// TIA Portal project "CraneSim" (V18)

(* hardware
DEVICE "S7-1500/ET200MP station_1"  S7-1500 station
   slot 0: "Rail_0"  Rack  6ES7 590-1***0-0AA0
   slot 1: "PLC_1"  CPU 1511-1 PN  6ES7 511-1AK02-0AB0  V2.9
      slot 3: "CPU display_1"  6ES7591-1AA00-0AA0
      slot 32768: "PROFINET interface_1"  X1
         slot 32769: "Port_1"  X1 P1
         slot 32770: "Port_2"  X1 P2
      slot 34817: "Virtual CP interface port_1"  Virtual CP interface port  Virtual CP interface port
*)

// ===== PLC "PLC_1"  CPU 1511-1 PN =====

VAR_GLOBAL   // PLC tag table "Default tag table"
   "Clock_Byte" AT %MB0 : Byte;
   "Clock_10Hz" AT %M0.0 : Bool;
   "Clock_5Hz" AT %M0.1 : Bool;
   "Clock_2.5Hz" AT %M0.2 : Bool;
   "Clock_2Hz" AT %M0.3 : Bool;
   "Clock_1.25Hz" AT %M0.4 : Bool;
   "Clock_1Hz" AT %M0.5 : Bool;
   "Clock_0.625Hz" AT %M0.6 : Bool;
   "Clock_0.5Hz" AT %M0.7 : Bool;
END_VAR

TYPE "typeTask"
   STRUCT
      station : Int;
      dwell_s : Int;
      crane : String[4];
      tank_name : String[10];
      prev : Int;
      next : Int;
      status : Int;
   END_STRUCT;
END_TYPE

DATA_BLOCK "Line4Data"   // DB2
{ S7_Optimized_Access := 'TRUE' }
VERSION : 0.1
   VAR
      task_count : Int;
      tasks : Array[1..20] of "typeTask";
      cmd_send : Bool;
      sts_busy : Bool;
      sts_done : Bool;
      sts_step : Int;
      sts_state : Int;
      ls_at : Array[0..9] of Bool;
      ls_dip : Bool;
      ls_up : Bool;
      btn_start : Bool;
      mv_fwd : Bool;
      mv_rev : Bool;
      mv_up : Bool;
      mv_down : Bool;
   END_VAR
BEGIN
END_DATA_BLOCK

DATA_BLOCK "CraneSequencer_DB"   // DB3
{ S7_Optimized_Access := 'TRUE' }
VERSION : 0.1
// stored: InstanceOfName CraneSequencer
"CraneSequencer"
BEGIN
END_DATA_BLOCK

FUNCTION_BLOCK "CraneSequencer"   // FB1, SCL
{ S7_Optimized_Access := 'TRUE' }
VERSION : 0.1
   VAR
      state : Int;
      idx : Int;
      count : Int;
      cur : Int;
      prevSend : Bool;
      tHold : TON_TIME;
      tDwell : TON_TIME;
   END_VAR
   VAR_TEMP
      target : Int;
      arrived : Bool;
   END_VAR
BEGIN
   // CraneSequencer — runs the Line4Data.tasks[] batch through the crane sequence.
   // Call every scan from OB1. Shared data lives in global DB "Line4Data".
   // Stations: 0=Parking 1=Loading 2..N=tanks.

   "Line4Data".sts_state := #state;

   CASE #state OF
       0:
           "Line4Data".mv_fwd := FALSE;
           "Line4Data".mv_rev := FALSE;
           "Line4Data".mv_up := FALSE;
           "Line4Data".mv_down := FALSE;
           "Line4Data".sts_busy := FALSE;
           "Line4Data".sts_step := 0;
           IF "Line4Data".cmd_send AND NOT #prevSend AND "Line4Data".task_count > 0 THEN
               #count := "Line4Data".task_count;
               #idx := 1;
               "Line4Data".sts_done := FALSE;
               "Line4Data".sts_busy := TRUE;
               #state := 10;
           END_IF;

       10:
           "Line4Data".sts_busy := TRUE;
           #target := 1;
           #arrived := "TravelTo"(target := #target, cur := #cur, atTarget := "Line4Data".ls_at[#target], fwd => "Line4Data".mv_fwd, rev => "Line4Data".mv_rev);
           IF #arrived THEN
               #cur := #target;
               "Line4Data".mv_fwd := FALSE;
               "Line4Data".mv_rev := FALSE;
               #state := 20;
           END_IF;

       20:
           "Line4Data".mv_up := FALSE;
           "Line4Data".mv_down := TRUE;
           IF "Line4Data".ls_dip THEN
               "Line4Data".mv_down := FALSE;
               #state := 30;
           END_IF;

       30:
           #tHold(IN := "Line4Data".btn_start,
                  PT := T#3S);
           IF #tHold.Q THEN
               #state := 40;
           END_IF;

       40:
           "Line4Data".mv_down := FALSE;
           "Line4Data".mv_up := TRUE;
           IF "Line4Data".ls_up THEN
               "Line4Data".mv_up := FALSE;
               #state := 50;
           END_IF;

       50:
           "Line4Data".sts_step := #idx;
           "Line4Data".tasks[#idx].status := 1;
           #target := "Line4Data".tasks[#idx].station;
           #arrived := "TravelTo"(target := #target, cur := #cur, atTarget := "Line4Data".ls_at[#target], fwd => "Line4Data".mv_fwd, rev => "Line4Data".mv_rev);
           IF #arrived THEN
               #cur := #target;
               "Line4Data".mv_fwd := FALSE;
               "Line4Data".mv_rev := FALSE;
               #state := 60;
           END_IF;

       60:
           "Line4Data".mv_up := FALSE;
           "Line4Data".mv_down := TRUE;
           IF "Line4Data".ls_dip THEN
               "Line4Data".mv_down := FALSE;
               #state := 70;
           END_IF;

       70:
           #tDwell(IN := TRUE,
                   PT := DINT_TO_TIME(INT_TO_DINT("Line4Data".tasks[#idx].dwell_s) * 1000));
           IF #tDwell.Q THEN
               #tDwell(IN := FALSE,
                       PT := T#0S);
               #state := 80;
           END_IF;

       80:
           "Line4Data".mv_down := FALSE;
           "Line4Data".mv_up := TRUE;
           IF "Line4Data".ls_up THEN
               "Line4Data".mv_up := FALSE;
               "Line4Data".tasks[#idx].status := 2;
               IF #idx < #count THEN
                   #idx := #idx + 1;
                   #state := 50;
               ELSE
                   #state := 85;
               END_IF;
           END_IF;

       85:
           #target := 0;
           #arrived := "TravelTo"(target := #target, cur := #cur, atTarget := "Line4Data".ls_at[#target], fwd => "Line4Data".mv_fwd, rev => "Line4Data".mv_rev);
           IF #arrived THEN
               #cur := #target;
               "Line4Data".mv_fwd := FALSE;
               "Line4Data".mv_rev := FALSE;
               #state := 90;
           END_IF;

       90:
           "Line4Data".sts_busy := FALSE;
           "Line4Data".sts_done := TRUE;
           IF NOT "Line4Data".cmd_send THEN
               "Line4Data".sts_done := FALSE;
               "Line4Data".sts_step := 0;
               #state := 0;
           END_IF;
   END_CASE;

   #prevSend := "Line4Data".cmd_send;
END_FUNCTION_BLOCK

FUNCTION "TravelTo" : Bool   // FC2, SCL
{ S7_Optimized_Access := 'TRUE' }
VERSION : 0.1
   VAR_INPUT
      target : Int;
      cur : Int;
      atTarget : Bool;
   END_VAR
   VAR_OUTPUT
      fwd : Bool;
      rev : Bool;
   END_VAR
BEGIN
   // TravelTo — pick the travel direction toward a target station.
   // Returns TRUE when the target limit switch is already made (arrived → stop).
   #fwd := FALSE;
   #rev := FALSE;

   IF #atTarget THEN
       ;                       // arrived: leave both motors off
   ELSIF #target > #cur THEN
       #fwd := TRUE;           // higher station number → travel forward
   ELSE
       #rev := TRUE;           // lower station number → travel reverse
   END_IF;

   #TravelTo := #atTarget;
END_FUNCTION

ORGANIZATION_BLOCK "Main"   // OB1, LAD, ProgramCycle
TITLE = "Main Program Sweep (Cycle)"
{ S7_Optimized_Access := 'TRUE' }
VERSION : 0.1
   VAR_INPUT
      Initial_Call : Bool;   // Initial call of this OB
      Remanence : Bool;   // =True, if remanent data are available
   END_VAR
BEGIN

REGION Network 1
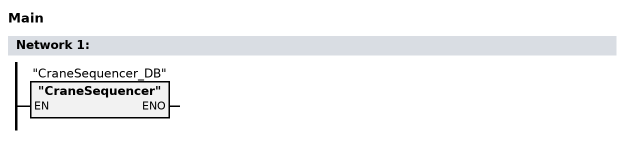
   RUNG wire#powerrail
      "CraneSequencer_DB"()
   END_RUNG
   // the same network as SCL:
   "CraneSequencer_DB"();   // "CraneSequencer"
END_REGION
END_ORGANIZATION_BLOCK